// TIA Portal project "Project4ă" (V18)

(* hardware
DEVICE "PC-System_1"  SIMATIC PC station
   slot 0: "SIMATIC PC station"  Rail  SIMATIC PC-Station  V1.0
      slot 125: "Stationmanager"  Station_Manager  V6.0.4
   slot 1: "HMI_RT_1"  WinCC RT Advanced  6AV2 104-0xxxx-xxxx  17.0.0.0
      slot 33792: "Computer interface"  Host interface
   slot 2: "IE general_1"  IE General  IE_CP  V8.2.0
      slot 1: "PROFINET interface"  IEGeneral.Interface.8.2.0
DEVICE "S7-300/ET200M station_1"  S7-300 station
   slot 0: "Rail_0"  Rail  6ES7 390-1***0-0AA0
   slot 2: "PLC_1"  CPU 314C-2 PN/DP  6ES7 314-6EH04-0AB0  V3.3.18
      slot 2: "PROFINET interface_1"  PN-IO
         slot 1: "Port_1"  Port
         slot 2: "Port_2"  Port
      slot 5: "DI 24/DO 16_1"  DI24/DO16
      slot 6: "AI 5/AO 2_1"  AI5/AO2
      slot 7: "Count_1"  Counter
      slot 8: "Positioning_1"  Positioning
*)

// ===== PLC "PLC_1"  CPU 314C-2 PN/DP =====

VAR_GLOBAL   // PLC tag table "Address"
   "START" AT %I0.0 : Bool;
   "S1" AT %I0.1 : Bool;
   "S2" AT %I0.2 : Bool;
   "S3" AT %I0.3 : Bool;
   "S4" AT %I0.4 : Bool;
   "SET" AT %I0.5 : Bool;
   "A+" AT %Q0.0 : Bool;
   "A-" AT %Q0.1 : Bool;
   "B+" AT %Q0.2 : Bool;
   "B-" AT %Q0.3 : Bool;
   "K1" AT %M0.0 : Bool;
   "K2" AT %M0.1 : Bool;
   "K3" AT %M0.2 : Bool;
   "K4" AT %M0.3 : Bool;
END_VAR

ORGANIZATION_BLOCK "Main"   // OB1, LAD
TITLE = "Main Program Sweep (Cycle)"
{ S7_Optimized_Access := 'FALSE' }
VERSION : 0.1
   VAR_TEMP
      OB1_EV_CLASS : Byte;   // Bits 0-3 = 1 (Coming event), Bits 4-7 = 1 (Event class 1)
      OB1_SCAN_1 : Byte;   // 1 (Cold restart scan 1 of OB 1), 3 (Scan 2-n of OB 1)
      OB1_PRIORITY : Byte;   // Priority of OB Execution
      OB1_OB_NUMBR : Byte;   // 1 (Organization block 1, OB1)
      OB1_RESERVED_1 : Byte;   // Reserved for system
      OB1_RESERVED_2 : Byte;   // Reserved for system
      OB1_PREV_CYCLE : Int;   // Cycle time of previous OB1 scan (milliseconds)
      OB1_MIN_CYCLE : Int;   // Minimum cycle time of OB1 (milliseconds)
      OB1_MAX_CYCLE : Int;   // Maximum cycle time of OB1 (milliseconds)
      OB1_DATE_TIME : Date_And_Time;   // Date and time OB1 started
   END_VAR
BEGIN

REGION Network 1: NHIP 1
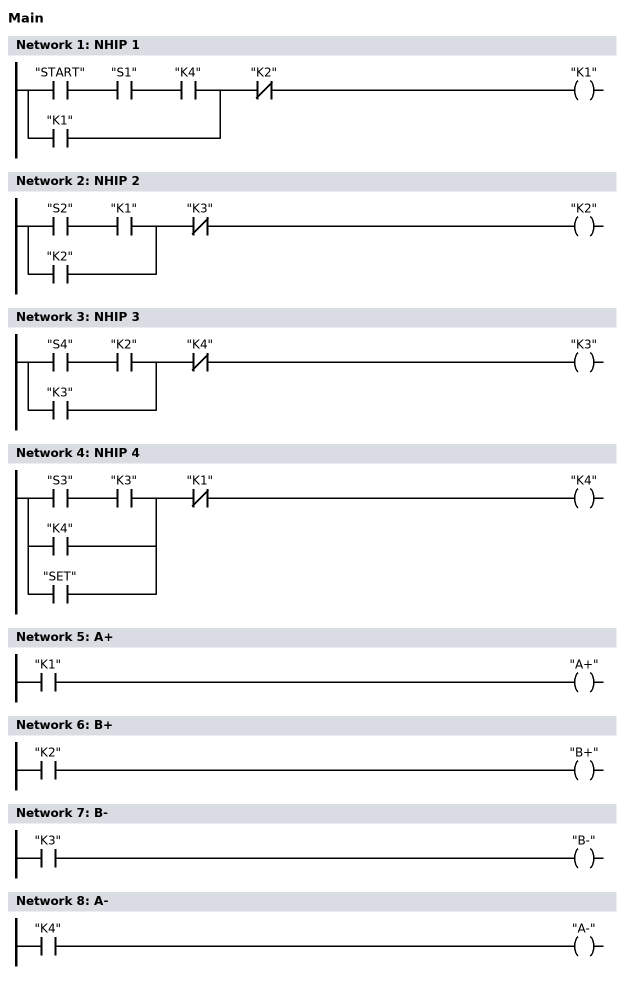
   RUNG wire#powerrail
      Contact( "START" )
      Contact( "S1" )
      Contact( "K4" )
      wire#w1
      I_Contact( "K2" )
      Coil( "K1" )
   END_RUNG
   RUNG wire#powerrail
      Contact( "K1" )
   END_RUNG wire#w1
   // the same network as SCL:
   "K1" := (("START" AND "S1" AND "K4") OR "K1") AND NOT "K2";
END_REGION

REGION Network 2: NHIP 2
   RUNG wire#powerrail
      Contact( "S2" )
      Contact( "K1" )
      wire#w1
      I_Contact( "K3" )
      Coil( "K2" )
   END_RUNG
   RUNG wire#powerrail
      Contact( "K2" )
   END_RUNG wire#w1
   // the same network as SCL:
   "K2" := (("S2" AND "K1") OR "K2") AND NOT "K3";
END_REGION

REGION Network 3: NHIP 3
   RUNG wire#powerrail
      Contact( "S4" )
      Contact( "K2" )
      wire#w1
      I_Contact( "K4" )
      Coil( "K3" )
   END_RUNG
   RUNG wire#powerrail
      Contact( "K3" )
   END_RUNG wire#w1
   // the same network as SCL:
   "K3" := (("S4" AND "K2") OR "K3") AND NOT "K4";
END_REGION

REGION Network 4: NHIP 4
   RUNG wire#powerrail
      Contact( "S3" )
      Contact( "K3" )
      wire#w1
      I_Contact( "K1" )
      Coil( "K4" )
   END_RUNG
   RUNG wire#powerrail
      Contact( "K4" )
   END_RUNG wire#w1
   RUNG wire#powerrail
      Contact( "SET" )
   END_RUNG wire#w1
   // the same network as SCL:
   "K4" := (("S3" AND "K3") OR "K4" OR "SET") AND NOT "K1";
END_REGION

REGION Network 5: A+
   RUNG wire#powerrail
      Contact( "K1" )
      Coil( "A+" )
   END_RUNG
   // the same network as SCL:
   "A+" := "K1";
END_REGION

REGION Network 6: B+
   RUNG wire#powerrail
      Contact( "K2" )
      Coil( "B+" )
   END_RUNG
   // the same network as SCL:
   "B+" := "K2";
END_REGION

REGION Network 7: B-
   RUNG wire#powerrail
      Contact( "K3" )
      Coil( "B-" )
   END_RUNG
   // the same network as SCL:
   "B-" := "K3";
END_REGION

REGION Network 8: A-
   RUNG wire#powerrail
      Contact( "K4" )
      Coil( "A-" )
   END_RUNG
   // the same network as SCL:
   "A-" := "K4";
END_REGION
END_ORGANIZATION_BLOCK

(* ===== HMI "HMI_RT_1" =====
connection "HMI_Connection_1": ETHERNET, S7_1200_OMS
connection "HMI_Connection_2": ETHERNET, S7_1200_OMS
*)